Fanuc KAREL source: KT00552.KL

PROGRAM KT00552
%NOLOCKGROUP
VAR
  P1: JOINTPOS
  P2: JOINTPOS
  OUT: JOINTPOS
BEGIN
  OUT = P1 : P2
END KT00552
